(* IEC 61131-3 sources: Godot-Digital-Twin/codesys/v1/pous, 6 files *)

(* ---- ST_DigitalTwinTCPConfiguration.st ---- *)
TYPE ST_DigitalTwinTCPConfiguration :
STRUCT
	sIpAddress	    : NBS.IPADDRESS := '127.0.0.1';
	uiPort		    : UINT		    := 50003;

	sDataHeader     : STRING	    := 'CRD';
	timSendDataTime : TIME 	        := T#10MS;
END_STRUCT
END_TYPE

(* ---- ST_DigitalTwinTCPData.st ---- *)
TYPE ST_DigitalTwinTCPData :
STRUCT
	uiNumberOfVariablesToSend		: UINT;
	arDataVariablesToSend			: ARRAY[1..GVL_DigitalTwinConstants.MaxNumberOfVariablesToSend] OF REAL;
END_STRUCT
END_TYPE

(* ---- GVL_DigitalTwinConstants.st ---- *)
{attribute 'qualified_only'}
VAR_GLOBAL CONSTANT
	MaxNumberOfVariablesToSend			: UINT := 10;
	ByteArraySize					    : UINT := 1024;

END_VAR

(* ---- FB_Clock.st ---- *)
FUNCTION_BLOCK FB_Clock
VAR_INPUT
	Enable : BOOL;
	Clock  : TIME;
END_VAR
VAR_OUTPUT
	Q      : BOOL;
END_VAR
VAR
	fbBlink : BLINK;
	fbRtrig : R_TRIG;
END_VAR

fbBlink(ENABLE:= Enable, TIMELOW:= Clock/2, TIMEHIGH:= Clock/2, OUT=> );
fbRtrig(CLK:= fbBlink.OUT, Q=> Q);

(* ---- FB_DigitalTwinTCPCommunication.st ---- *)
FUNCTION_BLOCK FB_DigitalTwinTCPCommunication
VAR_INPUT
	i_xEnable 	: BOOL;
END_VAR
VAR_OUTPUT
END_VAR
VAR
	fbTcpServer       : NBS.TCP_Server;
	fbTcpConnection   : NBS.TCP_Connection;
	fbSendDataClock	  : FB_Clock;
	fbIpAddress       : NBS.IPv4Address;
	xEnableConnection : BOOL;
	abSendData		  : ARRAY[1..GVL_DigitalTwinConstants.ByteArraySize] OF BYTE;
	udiSendDataSize	  : UDINT;
	iIndex			  : INT;

END_VAR

VAR_IN_OUT

	iq_stConfiguration : ST_DigitalTwinTCPConfiguration;
	iq_StData		   : ST_DigitalTwinTCPData;
END_VAR

IF fbTcpConnection._xSocketClosed THEN
	xEnableConnection := FALSE;

ELSIF i_xEnable THEN
	xEnableConnection := TRUE;

ELSE
	xEnableConnection := FALSE;

END_IF

IF fbIpAddress.ipAddress <> iq_stConfiguration.sIpAddress THEN
	fbIpAddress.SetInitialValue(ipAddress := iq_stConfiguration.sIpAddress);
END_IF

fbTcpServer(
	xEnable := i_xEnable,
    itfIPAddress := fbIpAddress,
    uiPort := iq_stConfiguration.uiPort );

fbTcpConnection(
	xEnable:= xEnableConnection,
     itfServer := fbTcpServer);

	 fbSendDataClock(Enable:= i_xEnable, Clock:= iq_stConfiguration.timSendDataTime, Q=> );

IF fbTcpConnection.xActive AND fbSendDataClock.Q THEN
	BuildSendData();
	fbTcpConnection.Write(pData := ADR(abSendData), udiSize := udiSendDataSize);
END_IF

// ===== BuildSendData =====
// Build the header

FOR iIndex := 1 TO Standard.LEN(iq_stConfiguration.sDataHeader) DO
	abSendData[iIndex] := iq_stConfiguration.sDataHeader[iIndex - 1];
END_FOR

// Number of variables - Byte

abSendData[Standard.LEN(iq_stConfiguration.sDataHeader) + 1] := UINT_TO_BYTE(iq_StData.uiNumberOfVariablesToSend);
MEMUtils.MemCpy(ADR(abSendData[Standard.LEN(iq_stConfiguration.sDataHeader)+ 2]) ,ADR(iq_StData.arDataVariablesToSend[1]),iq_stData.uiNumberOfVariablesToSend*4);
udiSendDataSize := INT_TO_UDINT(Standard.LEN(iq_stConfiguration.sDataHeader)) + 1 + iq_stData.uiNumberOfVariablesToSend*4;

(* ---- TCP_Communication.st ---- *)
PROGRAM TCP_Communication
VAR
	fbDigitalTwinTCPCommunication : FB_DigitalTwinTCPCommunication;
	fbDigitalTwinConfiguration    : ST_DigitalTwinTCPConfiguration;
	stDigitalTwinData			  : ST_DigitalTwinTCPData;
	xInitializationDone			  : BOOL;
END_VAR

IF NOT xInitializationDone THEN
	fbDigitalTwinConfiguration.sIpAddress      := '127.0.0.1';
	fbDigitalTwinConfiguration.uiPort          := 50003;
	fbDigitalTwinConfiguration.sDataHeader     := 'CRD';
	fbDigitalTwinConfiguration.timSendDataTime := T#10MS;

	xInitializationDone := TRUE;
END_IF

stDigitalTwinData.uiNumberOfVariablesToSend := 1;
stDigitalTwinData.arDataVariablesToSend[1] 	:= stDigitalTwinData.arDataVariablesToSend[1] + 1;

fbDigitalTwinTCPCommunication(i_xEnable:= TRUE, iq_stConfiguration:= fbDigitalTwinConfiguration, iq_StData:= stDigitalTwinData);
